Fanuc KAREL source: KT00469.KL

PROGRAM KT00469
%NOLOCKGROUP
VAR
  P1: JOINTPOS
  P2: XYZWPREXT
  OUT: BOOLEAN
BEGIN
    P2.Y = 2.0
  OUT = P1 >= P2
END KT00469
